FUNCTION_BLOCK ProjectInformation_Tests EXTENDS TcUnit.FB_TestSuite

Test_TitleAndCompany();
Test_VersionIsOnePointThree();

METHOD PRIVATE Test_TitleAndCompany
TcUnit.TEST(__POUNAME());

AssertEquals_WSTRING(Expected := "Intecre.File", Actual := Intecre_File.F_GetTitle(), Message := 'library title');
AssertEquals_WSTRING(Expected := "Intecre Ltd", Actual := Intecre_File.F_GetCompany(), Message := 'library company');

TEST_FINISHED_NAMED(__POUNAME());
END_METHOD

METHOD PRIVATE Test_VersionIsOnePointThree
VAR
  version : ST_LibVersion;
END_VAR
TcUnit.TEST(__POUNAME());

version := Intecre_File.F_GetVersion();
AssertEquals_STRING(Expected := '1.3.1.0', Actual := version.sVersion, Message := 'library version string');
AssertEquals_UINT(Expected := 1, Actual := version.iMajor, Message := 'major version');
AssertEquals_UINT(Expected := 3, Actual := version.iMinor, Message := 'minor version');

TEST_FINISHED_NAMED(__POUNAME());
END_METHOD

END_FUNCTION_BLOCK

(* stored: Version 1.1.0.1, ProductVersion 3.1.4026.19
   POU ProjectInformation_Tests: Id {381041a5-d514-4320-a47a-32ffbd50e26e}, SpecialFunc None
   Method Test_TitleAndCompany: Id {be2a7440-8e41-4f1a-82d3-867bafb63399}
   Method Test_VersionIsOnePointThree: Id {8b2c3e5b-555d-49f2-8762-cabcccde16ef} *)
